Fanuc KAREL source: kd00069.KL

-- PROVISIONAL review KL for V770-1; original PC SHA256 6eaa0cc4fcd46ff0d82cfe17461059b8ecbd8fd5b7c3c368bcb8421a0c0d3802
-- Incomplete behavior may be omitted. Consult companion uncertainty JSON. Do not deploy.
PROGRAM KD00069
%NOLOCKGROUP
VAR
  I : INTEGER
  J : INTEGER
  B : BOOLEAN
  R : REAL
  S : STRING[80]
BEGIN
  -- UNRESOLVED_PC offsets 5-18; opcodes 9D,81,18,9D,1B,9D,12,9C,13,04
  -- UNRESOLVED_PC offsets 23-27; opcodes 7F
END KD00069
